// TIA Portal project "conveyor_sorting_hmi" (V19)

(* hardware
DEVICE "S71500/ET200MP-Station_1"  S7-1500 station
   slot 0: "Profilschiene_0"  6ES7 590-1***0-0AA0
   slot 1: "PLC_1"  CPU 1511-1 PN  6ES7 511-1AK00-0AB0  V1.8
   slot 2: "AI 8xU/I/RTD/TC ST_1"  AI 8xU/I/RTD/TC ST  6ES7 531-7KF00-0AB0  V2.0
   slot 3: "AI 8xU/I/RTD/TC ST_2"  AI 8xU/I/RTD/TC ST  6ES7 531-7KF00-0AB0  V2.0
   slot 4: "AI 8xU/I/RTD/TC ST_3"  AI 8xU/I/RTD/TC ST  6ES7 531-7KF00-0AB0  V2.0
   slot 5: "AI 8xU/I/RTD/TC ST_4"  AI 8xU/I/RTD/TC ST  6ES7 531-7KF00-0AB0  V2.0
   slot 6: "DI 16x24VDC BA_1"  DI 16x24VDC BA  6ES7 521-1BH10-0AA0  V1.0
DEVICE "HMI_1"  KTP700 Basic PN
   slot 0: "HMI_1"  KTP700 Basic PN  6AV2 123-2GB03-0AX0  17.0.0.0
   slot 1: "HMI_RT_1"  KTP700 Basic PN  6AV2 123-2GB03-0AX0  17.0.0.0
   slot 5: "HMI_1.IE_CP_1"  PROFINET Interface  17.0.0.0
      slot 1: "PROFINET Interface_1"  PROFINET Interface
         slot 1: "Port_1"  Port
*)

// ===== PLC "PLC_1"  CPU 1511-1 PN =====

VAR_GLOBAL   // PLC tag table "Standard-Variablentabelle"
   "Tag_1" AT %E0.0 : Bool;
   "Tag_2" AT %A0.0 : Bool;
   "Tag_3" AT %E0.1 : Bool;
   "Tag_4" AT %I0.2 : Bool;
   "Tag_5" AT %I0.3 : Bool;
   "Tag_6" AT %Q0.1 : Bool;
   "Tag_7" AT %IW30 : Int;
   "Tag_8" AT %QW30 : Int;
   "Tag_9" AT %QW32 : Int;
END_VAR

DATA_BLOCK "DB_coveyorData"   // DB1
{ S7_Optimized_Access := 'TRUE' }
VERSION : 0.1
   VAR
      start_belt : Bool;
      stop_belt : Bool;
      reset_belt : Bool;
      belt_run : Bool;
      part_size_mm : Real;
      good_count : Int;
      reject_count : Int;
      batch_done : Int;
   END_VAR
BEGIN
END_DATA_BLOCK

DATA_BLOCK "FB_sorterLogic_DB"   // DB2
{ S7_Optimized_Access := 'TRUE' }
VERSION : 0.1
// stored: InstanceOfName FB_sorterLogic
"FB_sorterLogic"
BEGIN
END_DATA_BLOCK

DATA_BLOCK "FB_CONVEYORSIM_DB"   // DB3
{ S7_Optimized_Access := 'TRUE' }
VERSION : 0.1
// stored: InstanceOfName FB_CONVEYORSIM
"FB_CONVEYORSIM"
BEGIN
END_DATA_BLOCK

FUNCTION_BLOCK "FB_sorterLogic"   // FB1, SCL
{ S7_Optimized_Access := 'TRUE' }
VERSION : 0.1
BEGIN
   // Conveyor belt run/stop/reset, part size check (10.0..25.0 mm), and batch counter
   IF "DB_coveyorData".reset_belt THEN
       "DB_coveyorData".good_count := 0;
       "DB_coveyorData".reject_count := 0;
       "DB_coveyorData".batch_done := 0;
       "DB_coveyorData".belt_run := FALSE;
   END_IF;

   IF "DB_coveyorData".stop_belt THEN
       "DB_coveyorData".belt_run := FALSE;
   ELSIF "DB_coveyorData".start_belt THEN
       "DB_coveyorData".belt_run := TRUE;
   END_IF;

   IF "DB_coveyorData".belt_run AND ("DB_coveyorData".part_size_mm > 0.0) THEN
       IF ("DB_coveyorData".part_size_mm >= 10.0) AND ("DB_coveyorData".part_size_mm <= 25.0) THEN
           "DB_coveyorData".good_count := "DB_coveyorData".good_count + 1;
       ELSE
           "DB_coveyorData".reject_count := "DB_coveyorData".reject_count + 1;
       END_IF;

       // Reset part_size_mm after counting so one part isn't counted every scan
       "DB_coveyorData".part_size_mm := 0.0;
   END_IF;

   IF "DB_coveyorData".good_count >= 5 THEN
       "DB_coveyorData".batch_done := 1;
   ELSE
       "DB_coveyorData".batch_done := 0;
   END_IF;
END_FUNCTION_BLOCK

FUNCTION_BLOCK "FB_CONVEYORSIM"   // FB2, SCL
{ S7_Optimized_Access := 'TRUE' }
VERSION : 0.1
   VAR
      scan_timer : Int;
      send_reject : Bool;
   END_VAR
BEGIN
   // Simulates parts arriving every ~150 scans while belt_run is TRUE
   IF "DB_coveyorData".belt_run THEN
       #scan_timer := #scan_timer + 1;
       IF #scan_timer >= 150 THEN
           #scan_timer := 0;
           IF #send_reject THEN
               "DB_coveyorData".part_size_mm := 32.0; // Reject part (> 25.0 mm)
               #send_reject := FALSE;
           ELSE
               "DB_coveyorData".part_size_mm := 18.0; // Good part (10.0..25.0 mm)
               #send_reject := TRUE;
           END_IF;
       END_IF;
   ELSE
       #scan_timer := 0;
   END_IF;
END_FUNCTION_BLOCK

FUNCTION "MHJ-PLC-Lab-Function-S71500" : Void   // FC9000, SCL
{ S7_Optimized_Access := 'TRUE' }
VERSION : 0.1
   VAR_TEMP
      Value : Byte;
      ForCounter : Int;
   END_VAR
   VAR CONSTANT
      Value_01_DW : DWord := 16#1223_5486;
      Value_02_DW : DWord := 16#A6C9_D1F5;
   END_VAR
BEGIN

   #Value:=PEEK(area := 16#82,
        dbNumber := 0,
        byteOffset := 511);
   #Value := #Value + 1;

   POKE(area := 16#82,
        dbNumber := 0,
        byteOffset := 511,
        value := #Value);

   POKE(area := 16#82,
        dbNumber := 0,
        byteOffset := 1016,
        value := #Value_01_DW);
   POKE(area := 16#82,
        dbNumber := 0,
        byteOffset := 1020,
        value := #Value_02_DW);

   FOR #ForCounter := 0 TO 63 DO
       #Value:=PEEK(area := 16#1,
            dbNumber := 0,
            byteOffset := #ForCounter);
       POKE(area := 16#81,
            dbNumber := 0,
            byteOffset := #ForCounter,
            value := #Value);
   END_FOR;
   #Value := PEEK(area := 16#1,
                  dbNumber := 0,
                  byteOffset := 512);
   POKE(area := 16#82,
        dbNumber := 0,
        byteOffset := 512,
        value := #Value);
END_FUNCTION

ORGANIZATION_BLOCK "Main"   // OB1, FBD, ProgramCycle
TITLE = "Main Program Sweep (Cycle)"
{ S7_Optimized_Access := 'TRUE' }
VERSION : 0.1
   VAR_INPUT
      Initial_Call : Bool;   // Initial call of this OB
      Remanence : Bool;   // =True, if remanent data are available
   END_VAR
BEGIN

REGION Network 1
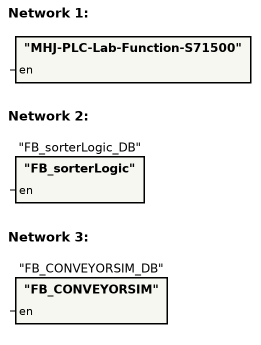
   "MHJ-PLC-Lab-Function-S71500"();
END_REGION

REGION Network 2
   "FB_sorterLogic_DB"();   // "FB_sorterLogic"
END_REGION

REGION Network 3
   "FB_CONVEYORSIM_DB"();   // "FB_CONVEYORSIM"
END_REGION
END_ORGANIZATION_BLOCK

(* ===== HMI "HMI_RT_1" =====
system functions are stored by id; their names below are inferred from use
connection "HMI_Connection_1": ETHERNET, SMART_S7_1500_OMS

HMI tags "Default tag table"
   "Tag_ScreenNumber" : UInt, internal
   "DB_coveyorData_start_belt" : Bool = PLC DB_coveyorData.start_belt, 1 s
   "DB_coveyorData_stop_belt" : Bool = PLC DB_coveyorData.stop_belt, 1 s
   "DB_coveyorData_reset_belt" : Bool = PLC DB_coveyorData.reset_belt, 1 s
   "DB_coveyorData_good_count" : Int = PLC DB_coveyorData.good_count, 1 s
   "DB_coveyorData_reject_count" : Int = PLC DB_coveyorData.reject_count, 1 s
   "DB_coveyorData_batch_done" : Int = PLC DB_coveyorData.batch_done, 1 s

Template "Template_1" 800x480
   Button "Exit" at 714,429 size 71x50; TextOff 'Exit'; PictureOff "ExitRuntime_KTP700_Basic_PN_TR"; PictureOn "ExitRuntime_KTP700_Basic_PN_TR"
      on Release: StopRuntime(0)
   Button "Template_Button" at 614,429 size 71x50; TextOff 'Text'
   Button "Template_Button_1" at 514,429 size 71x50; TextOff 'Text'
   Button "Template_Button_2" at 414,429 size 71x50; TextOff 'Text'
   Button "Template_Button_3" at 314,429 size 71x50; TextOff 'Text'
   Button "Template_Button_4" at 214,429 size 71x50; TextOff 'Text'
   Button "Alarms" at 114,429 size 71x50; TextOff 'Alarms'; PictureOff "AlarmDisplay_KTP700_Basic_PN_TR"; PictureOn "AlarmDisplay_KTP700_Basic_PN_TR"
      on Release: function_ef3f5d25("Alarm window_Unacknowledged", -1)
   Button "Start screen" at 14,429 size 71x50; TextOff 'Start screen'; PictureOff "NavigateHome_KTP700_Basic_PN_TR"; PictureOn "NavigateHome_KTP700_Basic_PN_TR"
      on Release: ActivateScreen("Root screen", 0)
   SymbolicIOField "Symbolic_IO_Field_Screen" at 93,9 size 600x33; TextOff '0'; TextOn '1'; TextList "TextList_ScreenNames"
      ProcessValue <- "Tag_ScreenNumber"
      on Change: ActivateScreenByNumber("Tag_ScreenNumber", 0)
   DateTimeField "HmiScreenItemData" at 695,25 size 105x25
   DateTimeField "HmiScreenItemData_1" at 695,0 size 105x25
   GraphicView "Logo" at 0,0 size 91x51; Picture "Logo of HMI_1"

screen "Root screen" 800x480, template "Template_1"
   on GenerateScreen: SetTag("Tag_ScreenNumber", 1)
   TextField "HmiScreenItemData" at 80,225 size 640x25; Text 'Welcome to HMI_1 (KTP700 Basic+ PN)!'
   Button "Button_1" at 54,90 size 96x32; TextOff 'start_belt'
      on Press: SetBit("DB_coveyorData_start_belt")
      on Release: ResetBit("DB_coveyorData_start_belt")
   Button "Button_2" at 195,90 size 96x32; TextOff 'stop_belt'
      on Press: SetBit("DB_coveyorData_stop_belt")
      on Release: ResetBit("DB_coveyorData_stop_belt")
   Button "Button_3" at 338,90 size 96x32; TextOff 'reset_bit'
      on Press: SetBit("DB_coveyorData_reset_belt")
      on Release: ResetBit("DB_coveyorData_reset_belt")
   IOField "I/O field_1" at 50,150 size 96x32; FormatPattern s999
      ProcessValue <- "DB_coveyorData_good_count"
   IOField "I/O field_2" at 187,150 size 96x32; FormatPattern s999
      ProcessValue <- "DB_coveyorData_reject_count"
   IOField "I/O field_3" at 332,150 size 96x32; FormatPattern s999
      ProcessValue <- "DB_coveyorData_batch_done"
*)